(* IEC 61131-3 sources: Test-Git_ESME26/TestProgettoESME_26.fbsproj/TemplateFullProgrammingFramework_Migration.device.xml.v3^/Plc Logic.plclogic.xml.v3^/Application.application.xml.v3^/TemplateFullProgrammingFramework/Tools, 2 files *)

(* ---- FC_IsDriveVirtual.fn.st ---- *)
FUNCTION FC_IsDriveVirtual : BOOL
VAR_INPUT
	i_ifDrive	: MOIN.IF_Axis;
END_VAR

VAR_OUTPUT
	q_etDiag	: GD.ET_Diag := GD.ET_Diag.Ok;
	q_etDiagExt	: ET_DiagExt := ET_DiagExt.Ok;
	q_sMsg		: STRING[80];
END_VAR

VAR
	xSuccess			: BOOL;
	ifWorkingModeAccess :  CFDI.IF_WorkingModeAccess;
	ifGetParentDevice   : DTSI.IF_GetParentDevice;
	ifDeviceAccess		: DTSI.IF_DeviceAccess;
END_VAR

IF i_ifDrive = 0 THEN
	q_etDiag	:= GD.ET_Diag.InputParameterInvalid;
	q_etDiagExt	:= ET_DiagExt.DriveInvalid;
	q_sMsg		:= 'FC_IsDriveVirtual: i_ifDrive not set';
ELSE
	xSuccess := __QUERYINTERFACE(i_ifDrive, ifGetParentDevice);
	IF NOT xSuccess OR ifGetParentDevice = 0 THEN
		// not a device-tree axis with user functions -> virtual axis
		FC_IsDriveVirtual := TRUE;
		RETURN;
	END_IF
	ifDeviceAccess := ifGetParentDevice.GetParentDevice();

	xSuccess := __QUERYINTERFACE(ifDeviceAccess, ifWorkingModeAccess);
	IF NOT xSuccess OR ifWorkingModeAccess = 0 THEN
		// not a device-tree axis with user functions -> virtual axis
		FC_IsDriveVirtual := TRUE;
	ELSE
		// device-tree axis with user funciton working mode -> read out working mode
		FC_IsDriveVirtual := (ifWorkingModeAccess.WorkingMode.DesiredMode = CFDI.ET_WorkingMode.Virtual);
	END_IF
END_IF

(* ---- FC_SetDeadTimeCompensation.fn.st ---- *)
FUNCTION FC_SetDeadTimeCompensation : BOOL
VAR_INPUT
	i_stSubModuleInterfaceMain		: AXM_ST_Main;
END_VAR
VAR
(* Init related variables *)
	//stLogicalAddressMaster			: SystemConfigurationItf.ST_LogicalAddress;
	lrShaftRefDelay					: LREAL;
	lrPositionDelay					: LREAL;
	diResult						: DINT;

END_VAR

(*
IF i_stSubModuleInterfaceMain.i_ifMaster <> 0 AND i_stSubModuleInterfaceMain.i_ifDrive <> 0 THEN
	stLogicalAddressMaster := i_stSubModuleInterfaceMain.i_ifMaster.stLogicalAddress;
	IF (stLogicalAddressMaster.udiType = SYSTEMINTERFACE.P_ENC_TYPE.udiType) OR			(* Physical encoder *)
		(stLogicalAddressMaster.udiType = SYSTEMINTERFACE.INC_IN_TYPE.udiType) OR		(* Incremental	encoder *)
		(stLogicalAddressMaster.udiType = SYSTEMINTERFACE.V_ENC_TYPE.udiType) THEN		(* Virtual master encoder *)

		stLogicalAddressMaster := i_stSubModuleInterfaceMain.i_ifDrive.stLogicalAddress;
		stLogicalAddressMaster.udiParameterId := 16#00A2;
		diResult := SYSTEMINTERFACE.FC_GetParameter(i_stLogAdr	:= stLogicalAddressMaster,
													i_dwBuffer	:= ADR(lrShaftRefDelay),
													i_diSize	:= SIZEOF(lrShaftRefDelay));
		IF diResult = 0 THEN
			i_stSubModuleInterfaceMain.iq_lencEncoder.Delay := -lrShaftRefDelay;
		END_IF
	ELSIF (stLogicalAddressMaster.udiType = SYSTEMINTERFACE.INC_IN3_TYPE.udiType) THEN  (* IncIn via TM5 TM5SE1IC20005 *)
		stLogicalAddressMaster := i_stSubModuleInterfaceMain.i_ifDrive.stLogicalAddress;
		stLogicalAddressMaster.udiParameterId := 16#00A2;
		diResult := SYSTEMINTERFACE.FC_GetParameter(i_stLogAdr	:= stLogicalAddressMaster,
													i_dwBuffer	:= ADR(lrShaftRefDelay),
													i_diSize	:= SIZEOF(lrShaftRefDelay));
		IF diResult = 0 THEN
			i_stSubModuleInterfaceMain.iq_lencEncoder.Delay := -lrShaftRefDelay;
			stLogicalAddressMaster := i_stSubModuleInterfaceMain.i_ifMaster.stLogicalAddress;
			stLogicalAddressMaster.udiParameterId := 16#008E; 					(* Parameter PositionDelay of TM5SE1IC20005 *)
			diResult := SYSTEMINTERFACE.FC_GetParameter(i_stLogAdr	:= stLogicalAddressMaster,
														i_dwBuffer	:= ADR(lrPositionDelay),
														i_diSize	:= SIZEOF(lrPositionDelay));
			IF diResult = 0 THEN
				i_stSubModuleInterfaceMain.iq_lencEncoder.Delay := -(lrShaftRefDelay + (-lrPositionDelay)) ;
			END_IF
		END_IF
	END_IF
END_IF
*)
IF diResult = 0 THEN
	FC_SetDeadTimeCompensation := TRUE;
END_IF
